// LS Electric XG5000 project: motor-control
// PLC LSPLC

PROGRAM motor_control (task: 스캔 프로그램)

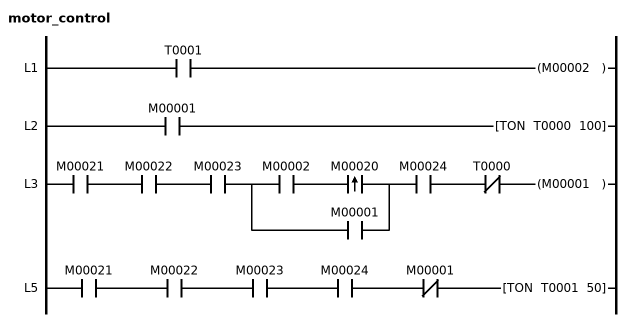
; L1
LOAD      T0001
OUT       M00002
; L2
LOAD      M00001
TON       T0000 100
; L3
LOAD      M00021
AND       M00022
AND       M00023
LOAD      M00002
ANDP      M00020
OR        M00001
AND LOAD
AND       M00024
AND NOT   T0000
OUT       M00001
; L5
LOAD      M00021
AND       M00022
AND       M00023
AND       M00024
AND NOT   M00001
TON       T0001 50